(* IEC 61131-3 sources: plc-st-coding-agent/progress/evidence/f14_v14_remaining_20261113/jobs/custom_minimax-m27 (part 5) *)

(* ---- public-medium-05.candidate_04.st ---- *)
(* ENGINEERING_CONTRACT
 * =============================================================================
 * Mode Switching (PUB001): Mode=0 manual, Mode=1 automatic. Output state on
 *   mode transition: both Motor outputs cleared, CompletionLight cleared.
 *   Transition detected via rising edge on Mode input variable.
 * Manual Mode (PUB002/PUB003):
 *   - Activation: Mode=0
 *   - Retention: MotorForward holds while ForwardButton=1 AND ReverseButton=0
 *   - Retention: MotorReverse holds while ReverseButton=1 AND ForwardButton=0
 *   - Deactivation: both cleared on any of: ForwardButton=0, ReverseButton=0,
 *     forward+reverse both asserted (interlock drops both), or Mode→1
 *   - Units: combinational, no timer
 * Automatic Mode (PUB004-PUB008):
 *   - Scan behavior: edge-sensitive state machine evaluated every scan
 *   - STATION_A activation: SensorA=TRUE AND State=IDLE
 *   - STATION_B activation: SensorB=TRUE AND State=MOVING_TO_B
 *   - STATION_C activation: SensorC=TRUE AND State=MOVING_TO_C
 *   - MotorForward activation: (State=IDLE AND SensorA=TRUE→ButtonA=TRUE)
 *     OR (State=STATION_A AND ButtonA=TRUE) OR (State=STATION_B AND ButtonB=TRUE)
 *   - MotorForward deactivation: on SensorB (→STATION_B) or SensorC (→STATION_C)
 *   - CompletionLight activation: SensorC=TRUE AND ButtonC=TRUE AND State=STATION_C
 *   - CompletionLight retention: holds until SensorC=FALSE (product removed)
 *   - CompletionLight deactivation: SensorC=FALSE transitions to IDLE
 *   - IDLE reset: State=IDLE when no product detected at any station
 *   - Units: boolean states, no timers
 * Same-scan priority: manual overrides automatic (Mode check first). Within
 *   automatic, state transition clears prior MotorForward before next sensor
 *   evaluation; CompletionLight set after Mode/state checks finalized.
 * Physical interlock: Pub002 prohibits MotorForward AND MotorReverse together.
 * =============================================================================
 *)

(* CONTRACT_RULES [] *)

FUNCTION_BLOCK ProductionLineControl
VAR_INPUT
    Mode            : BOOL;  (* 0=manual, 1=automatic *)
    ForwardButton   : BOOL;
    ReverseButton   : BOOL;
    SensorA         : BOOL;
    SensorB         : BOOL;
    SensorC         : BOOL;
    ButtonA         : BOOL;
    ButtonB         : BOOL;
    ButtonC         : BOOL;
END_VAR
VAR_OUTPUT
    MotorForward    : BOOL;
    MotorReverse    : BOOL;
    CompletionLight : BOOL;
END_VAR
VAR_CONSTANT
    IDLE         : INT := 0;
    STATION_A    : INT := 1;
    MOVING_TO_B  : INT := 2;
    STATION_B    : INT := 3;
    MOVING_TO_C  : INT := 4;
    STATION_C    : INT := 5;
END_VAR_CONSTANT

VAR
    State           : INT;  (* 0=IDLE, 1=STATION_A, 2=MOVING_TO_B, 3=STATION_B,
                                4=MOVING_TO_C, 5=STATION_C *)
    tmp_PreviousMode : BOOL;
    tmp_ModeRising   : BOOL;
END_VAR

    (* Constants for state identification *)
    (* Detect mode transition for reset behavior *)
    tmp_ModeRising := Mode AND NOT tmp_PreviousMode;
    tmp_PreviousMode := Mode;

    (* Reset outputs on mode entry into automatic *)
    IF tmp_ModeRising THEN
        MotorForward    := FALSE;
        MotorReverse    := FALSE;
        CompletionLight := FALSE;
    END_IF;

    (* Mode-based operation dispatch *)
    IF Mode = FALSE THEN
        (* Manual Mode (PUB002/PUB003) *)
        (* Interlock: forward and reverse cannot be energized together *)
        IF ForwardButton AND NOT ReverseButton THEN
            MotorForward := TRUE;
            MotorReverse := FALSE;
        ELSIF ReverseButton AND NOT ForwardButton THEN
            MotorForward := FALSE;
            MotorReverse := TRUE;
        ELSE
            MotorForward := FALSE;
            MotorReverse := FALSE;
        END_IF;
    ELSE
        (* Automatic Mode (PUB004-PUB008) *)
        MotorForward    := FALSE;
        MotorReverse    := FALSE;

        (* State machine evaluation *)
        CASE State OF
            IDLE :
                (* Wait for product at Workstation A *)
                IF SensorA THEN
                    State := STATION_A;
                END_IF;

            STATION_A :
                (* Product at Workstation A, wait for ButtonA *)
                IF ButtonA THEN
                    MotorForward := TRUE;
                    State := MOVING_TO_B;
                END_IF;
                (* Fallback: if product leaves A unexpectedly, return to IDLE *)
                IF NOT SensorA THEN
                    State := IDLE;
                END_IF;

            MOVING_TO_B :
                (* Motor running forward, wait for SensorB *)
                MotorForward := TRUE;
                IF SensorB THEN
                    MotorForward := FALSE;
                    State := STATION_B;
                END_IF;

            STATION_B :
                (* Product at Workstation B, wait for ButtonB *)
                IF ButtonB THEN
                    MotorForward := TRUE;
                    State := MOVING_TO_C;
                END_IF;
                (* Fallback: if product leaves B unexpectedly, return to IDLE *)
                IF NOT SensorB THEN
                    State := IDLE;
                END_IF;

            MOVING_TO_C :
                (* Motor running forward, wait for SensorC *)
                MotorForward := TRUE;
                IF SensorC THEN
                    MotorForward := FALSE;
                    State := STATION_C;
                END_IF;

            STATION_C :
                (* Product at Workstation C, wait for ButtonC, then product removal *)
                IF ButtonC THEN
                    CompletionLight := TRUE;
                END_IF;
                (* Product taken away: light off, return to IDLE *)
                IF NOT SensorC THEN
                    CompletionLight := FALSE;
                    State := IDLE;
                END_IF;

        END_CASE;
    END_IF;

END_FUNCTION_BLOCK

(* ---- public-medium-05.patch_base_02.st ---- *)
(* ENGINEERING_CONTRACT
 * =============================================================================
 * Mode Switching (PUB001): Mode=0 manual, Mode=1 automatic. Output state on
 *   mode transition: both Motor outputs cleared, CompletionLight cleared.
 *   Transition detected via rising edge on Mode input variable.
 * Manual Mode (PUB002/PUB003):
 *   - Activation: Mode=0
 *   - Retention: MotorForward holds while ForwardButton=1 AND ReverseButton=0
 *   - Retention: MotorReverse holds while ReverseButton=1 AND ForwardButton=0
 *   - Deactivation: both cleared on any of: ForwardButton=0, ReverseButton=0,
 *     forward+reverse both asserted (interlock drops both), or Mode→1
 *   - Units: combinational, no timer
 * Automatic Mode (PUB004-PUB008):
 *   - Scan behavior: edge-sensitive state machine evaluated every scan
 *   - STATION_A activation: SensorA=TRUE AND State=IDLE
 *   - STATION_B activation: SensorB=TRUE AND State=MOVING_TO_B
 *   - STATION_C activation: SensorC=TRUE AND State=MOVING_TO_C
 *   - MotorForward activation: (State=IDLE AND SensorA=TRUE→ButtonA=TRUE)
 *     OR (State=STATION_A AND ButtonA=TRUE) OR (State=STATION_B AND ButtonB=TRUE)
 *   - MotorForward deactivation: on SensorB (→STATION_B) or SensorC (→STATION_C)
 *   - CompletionLight activation: SensorC=TRUE AND ButtonC=TRUE AND State=STATION_C
 *   - CompletionLight retention: holds until SensorC=FALSE (product removed)
 *   - CompletionLight deactivation: SensorC=FALSE transitions to IDLE
 *   - IDLE reset: State=IDLE when no product detected at any station
 *   - Units: boolean states, no timers
 * Same-scan priority: manual overrides automatic (Mode check first). Within
 *   automatic, state transition clears prior MotorForward before next sensor
 *   evaluation; CompletionLight set after Mode/state checks finalized.
 * Physical interlock: Pub002 prohibits MotorForward AND MotorReverse together.
 * =============================================================================
 *)

(* CONTRACT_RULES [] *)

FUNCTION_BLOCK ProductionLineControl
VAR_INPUT
    Mode            : BOOL;  (* 0=manual, 1=automatic *)
    ForwardButton   : BOOL;
    ReverseButton   : BOOL;
    SensorA         : BOOL;
    SensorB         : BOOL;
    SensorC         : BOOL;
    ButtonA         : BOOL;
    ButtonB         : BOOL;
    ButtonC         : BOOL;
END_VAR
VAR_OUTPUT
    MotorForward    : BOOL;
    MotorReverse    : BOOL;
    CompletionLight : BOOL;
END_VAR
VAR
    State           : INT;  (* 0=IDLE, 1=STATION_A, 2=MOVING_TO_B, 3=STATION_B,
                                4=MOVING_TO_C, 5=STATION_C *)
    tmp_PreviousMode : BOOL;
    tmp_ModeRising   : BOOL;
END_VAR

    (* Constants for state identification *)
    CONST
        IDLE         : INT := 0;
        STATION_A    : INT := 1;
        MOVING_TO_B  : INT := 2;
        STATION_B    : INT := 3;
        MOVING_TO_C  : INT := 4;
        STATION_C    : INT := 5;
    END_CONST

    (* Detect mode transition for reset behavior *)
    tmp_ModeRising := Mode AND NOT tmp_PreviousMode;
    tmp_PreviousMode := Mode;

    (* Reset outputs on mode entry into automatic *)
    IF tmp_ModeRising THEN
        MotorForward    := FALSE;
        MotorReverse    := FALSE;
        CompletionLight := FALSE;
    END_IF;

    (* Mode-based operation dispatch *)
    IF Mode = FALSE THEN
        (* Manual Mode (PUB002/PUB003) *)
        (* Interlock: forward and reverse cannot be energized together *)
        IF ForwardButton AND NOT ReverseButton THEN
            MotorForward := TRUE;
            MotorReverse := FALSE;
        ELSIF ReverseButton AND NOT ForwardButton THEN
            MotorForward := FALSE;
            MotorReverse := TRUE;
        ELSE
            MotorForward := FALSE;
            MotorReverse := FALSE;
        END_IF;
    ELSE
        (* Automatic Mode (PUB004-PUB008) *)
        MotorForward    := FALSE;
        MotorReverse    := FALSE;

        (* State machine evaluation *)
        CASE State OF
            IDLE :
                (* Wait for product at Workstation A *)
                IF SensorA THEN
                    State := STATION_A;
                END_IF;

            STATION_A :
                (* Product at Workstation A, wait for ButtonA *)
                IF ButtonA THEN
                    MotorForward := TRUE;
                    State := MOVING_TO_B;
                END_IF;
                (* Fallback: if product leaves A unexpectedly, return to IDLE *)
                IF NOT SensorA THEN
                    State := IDLE;
                END_IF;

            MOVING_TO_B :
                (* Motor running forward, wait for SensorB *)
                MotorForward := TRUE;
                IF SensorB THEN
                    MotorForward := FALSE;
                    State := STATION_B;
                END_IF;

            STATION_B :
                (* Product at Workstation B, wait for ButtonB *)
                IF ButtonB THEN
                    MotorForward := TRUE;
                    State := MOVING_TO_C;
                END_IF;
                (* Fallback: if product leaves B unexpectedly, return to IDLE *)
                IF NOT SensorB THEN
                    State := IDLE;
                END_IF;

            MOVING_TO_C :
                (* Motor running forward, wait for SensorC *)
                MotorForward := TRUE;
                IF SensorC THEN
                    MotorForward := FALSE;
                    State := STATION_C;
                END_IF;

            STATION_C :
                (* Product at Workstation C, wait for ButtonC, then product removal *)
                IF ButtonC THEN
                    CompletionLight := TRUE;
                END_IF;
                (* Product taken away: light off, return to IDLE *)
                IF NOT SensorC THEN
                    CompletionLight := FALSE;
                    State := IDLE;
                END_IF;

        END_CASE;
    END_IF;

END_FUNCTION_BLOCK

(* ---- public-medium-05.patch_base_03.st ---- *)
TYPE ProductionState : INT (
    IDLE := 0,
    STATION_A := 1,
    MOVING_TO_B := 2,
    STATION_B := 3,
    MOVING_TO_C := 4,
    STATION_C := 5
);
END_TYPE;

(* ENGINEERING_CONTRACT
 * =============================================================================
 * Mode Switching (PUB001): Mode=0 manual, Mode=1 automatic. Output state on
 *   mode transition: both Motor outputs cleared, CompletionLight cleared.
 *   Transition detected via rising edge on Mode input variable.
 * Manual Mode (PUB002/PUB003):
 *   - Activation: Mode=0
 *   - Retention: MotorForward holds while ForwardButton=1 AND ReverseButton=0
 *   - Retention: MotorReverse holds while ReverseButton=1 AND ForwardButton=0
 *   - Deactivation: both cleared on any of: ForwardButton=0, ReverseButton=0,
 *     forward+reverse both asserted (interlock drops both), or Mode→1
 *   - Units: combinational, no timer
 * Automatic Mode (PUB004-PUB008):
 *   - Scan behavior: edge-sensitive state machine evaluated every scan
 *   - STATION_A activation: SensorA=TRUE AND State=IDLE
 *   - STATION_B activation: SensorB=TRUE AND State=MOVING_TO_B
 *   - STATION_C activation: SensorC=TRUE AND State=MOVING_TO_C
 *   - MotorForward activation: (State=IDLE AND SensorA=TRUE→ButtonA=TRUE)
 *     OR (State=STATION_A AND ButtonA=TRUE) OR (State=STATION_B AND ButtonB=TRUE)
 *   - MotorForward deactivation: on SensorB (→STATION_B) or SensorC (→STATION_C)
 *   - CompletionLight activation: SensorC=TRUE AND ButtonC=TRUE AND State=STATION_C
 *   - CompletionLight retention: holds until SensorC=FALSE (product removed)
 *   - CompletionLight deactivation: SensorC=FALSE transitions to IDLE
 *   - IDLE reset: State=IDLE when no product detected at any station
 *   - Units: boolean states, no timers
 * Same-scan priority: manual overrides automatic (Mode check first). Within
 *   automatic, state transition clears prior MotorForward before next sensor
 *   evaluation; CompletionLight set after Mode/state checks finalized.
 * Physical interlock: Pub002 prohibits MotorForward AND MotorReverse together.
 * =============================================================================
 *)

(* CONTRACT_RULES [] *)

FUNCTION_BLOCK ProductionLineControl
VAR_INPUT
    Mode            : BOOL;  (* 0=manual, 1=automatic *)
    ForwardButton   : BOOL;
    ReverseButton   : BOOL;
    SensorA         : BOOL;
    SensorB         : BOOL;
    SensorC         : BOOL;
    ButtonA         : BOOL;
    ButtonB         : BOOL;
    ButtonC         : BOOL;
END_VAR
VAR_OUTPUT
    MotorForward    : BOOL;
    MotorReverse    : BOOL;
    CompletionLight : BOOL;
END_VAR
VAR
    State           : INT;  (* 0=IDLE, 1=STATION_A, 2=MOVING_TO_B, 3=STATION_B,
                                4=MOVING_TO_C, 5=STATION_C *)
    tmp_PreviousMode : BOOL;
    tmp_ModeRising   : BOOL;
END_VAR

    (* Constants for state identification *)
    (* Detect mode transition for reset behavior *)
    tmp_ModeRising := Mode AND NOT tmp_PreviousMode;
    tmp_PreviousMode := Mode;

    (* Reset outputs on mode entry into automatic *)
    IF tmp_ModeRising THEN
        MotorForward    := FALSE;
        MotorReverse    := FALSE;
        CompletionLight := FALSE;
    END_IF;

    (* Mode-based operation dispatch *)
    IF Mode = FALSE THEN
        (* Manual Mode (PUB002/PUB003) *)
        (* Interlock: forward and reverse cannot be energized together *)
        IF ForwardButton AND NOT ReverseButton THEN
            MotorForward := TRUE;
            MotorReverse := FALSE;
        ELSIF ReverseButton AND NOT ForwardButton THEN
            MotorForward := FALSE;
            MotorReverse := TRUE;
        ELSE
            MotorForward := FALSE;
            MotorReverse := FALSE;
        END_IF;
    ELSE
        (* Automatic Mode (PUB004-PUB008) *)
        MotorForward    := FALSE;
        MotorReverse    := FALSE;

        (* State machine evaluation *)
        CASE State OF
            IDLE :
                (* Wait for product at Workstation A *)
                IF SensorA THEN
                    State := STATION_A;
                END_IF;

            STATION_A :
                (* Product at Workstation A, wait for ButtonA *)
                IF ButtonA THEN
                    MotorForward := TRUE;
                    State := MOVING_TO_B;
                END_IF;
                (* Fallback: if product leaves A unexpectedly, return to IDLE *)
                IF NOT SensorA THEN
                    State := IDLE;
                END_IF;

            MOVING_TO_B :
                (* Motor running forward, wait for SensorB *)
                MotorForward := TRUE;
                IF SensorB THEN
                    MotorForward := FALSE;
                    State := STATION_B;
                END_IF;

            STATION_B :
                (* Product at Workstation B, wait for ButtonB *)
                IF ButtonB THEN
                    MotorForward := TRUE;
                    State := MOVING_TO_C;
                END_IF;
                (* Fallback: if product leaves B unexpectedly, return to IDLE *)
                IF NOT SensorB THEN
                    State := IDLE;
                END_IF;

            MOVING_TO_C :
                (* Motor running forward, wait for SensorC *)
                MotorForward := TRUE;
                IF SensorC THEN
                    MotorForward := FALSE;
                    State := STATION_C;
                END_IF;

            STATION_C :
                (* Product at Workstation C, wait for ButtonC, then product removal *)
                IF ButtonC THEN
                    CompletionLight := TRUE;
                END_IF;
                (* Product taken away: light off, return to IDLE *)
                IF NOT SensorC THEN
                    CompletionLight := FALSE;
                    State := IDLE;
                END_IF;

        END_CASE;
    END_IF;

END_FUNCTION_BLOCK

(* ---- public-medium-05.patch_base_04.st ---- *)
CONST
    IDLE         : INT := 0;
    STATION_A    : INT := 1;
    MOVING_TO_B  : INT := 2;
    STATION_B    : INT := 3;
    MOVING_TO_C  : INT := 4;
    STATION_C    : INT := 5;
END_CONST

(* ENGINEERING_CONTRACT
 * =============================================================================
 * Mode Switching (PUB001): Mode=0 manual, Mode=1 automatic. Output state on
 *   mode transition: both Motor outputs cleared, CompletionLight cleared.
 *   Transition detected via rising edge on Mode input variable.
 * Manual Mode (PUB002/PUB003):
 *   - Activation: Mode=0
 *   - Retention: MotorForward holds while ForwardButton=1 AND ReverseButton=0
 *   - Retention: MotorReverse holds while ReverseButton=1 AND ForwardButton=0
 *   - Deactivation: both cleared on any of: ForwardButton=0, ReverseButton=0,
 *     forward+reverse both asserted (interlock drops both), or Mode→1
 *   - Units: combinational, no timer
 * Automatic Mode (PUB004-PUB008):
 *   - Scan behavior: edge-sensitive state machine evaluated every scan
 *   - STATION_A activation: SensorA=TRUE AND State=IDLE
 *   - STATION_B activation: SensorB=TRUE AND State=MOVING_TO_B
 *   - STATION_C activation: SensorC=TRUE AND State=MOVING_TO_C
 *   - MotorForward activation: (State=IDLE AND SensorA=TRUE→ButtonA=TRUE)
 *     OR (State=STATION_A AND ButtonA=TRUE) OR (State=STATION_B AND ButtonB=TRUE)
 *   - MotorForward deactivation: on SensorB (→STATION_B) or SensorC (→STATION_C)
 *   - CompletionLight activation: SensorC=TRUE AND ButtonC=TRUE AND State=STATION_C
 *   - CompletionLight retention: holds until SensorC=FALSE (product removed)
 *   - CompletionLight deactivation: SensorC=FALSE transitions to IDLE
 *   - IDLE reset: State=IDLE when no product detected at any station
 *   - Units: boolean states, no timers
 * Same-scan priority: manual overrides automatic (Mode check first). Within
 *   automatic, state transition clears prior MotorForward before next sensor
 *   evaluation; CompletionLight set after Mode/state checks finalized.
 * Physical interlock: Pub002 prohibits MotorForward AND MotorReverse together.
 * =============================================================================
 *)

(* CONTRACT_RULES [] *)

FUNCTION_BLOCK ProductionLineControl
VAR_INPUT
    Mode            : BOOL;  (* 0=manual, 1=automatic *)
    ForwardButton   : BOOL;
    ReverseButton   : BOOL;
    SensorA         : BOOL;
    SensorB         : BOOL;
    SensorC         : BOOL;
    ButtonA         : BOOL;
    ButtonB         : BOOL;
    ButtonC         : BOOL;
END_VAR
VAR_OUTPUT
    MotorForward    : BOOL;
    MotorReverse    : BOOL;
    CompletionLight : BOOL;
END_VAR
VAR
    State           : INT;  (* 0=IDLE, 1=STATION_A, 2=MOVING_TO_B, 3=STATION_B,
                                4=MOVING_TO_C, 5=STATION_C *)
    tmp_PreviousMode : BOOL;
    tmp_ModeRising   : BOOL;
END_VAR

    (* Constants for state identification *)
    (* Detect mode transition for reset behavior *)
    tmp_ModeRising := Mode AND NOT tmp_PreviousMode;
    tmp_PreviousMode := Mode;

    (* Reset outputs on mode entry into automatic *)
    IF tmp_ModeRising THEN
        MotorForward    := FALSE;
        MotorReverse    := FALSE;
        CompletionLight := FALSE;
    END_IF;

    (* Mode-based operation dispatch *)
    IF Mode = FALSE THEN
        (* Manual Mode (PUB002/PUB003) *)
        (* Interlock: forward and reverse cannot be energized together *)
        IF ForwardButton AND NOT ReverseButton THEN
            MotorForward := TRUE;
            MotorReverse := FALSE;
        ELSIF ReverseButton AND NOT ForwardButton THEN
            MotorForward := FALSE;
            MotorReverse := TRUE;
        ELSE
            MotorForward := FALSE;
            MotorReverse := FALSE;
        END_IF;
    ELSE
        (* Automatic Mode (PUB004-PUB008) *)
        MotorForward    := FALSE;
        MotorReverse    := FALSE;

        (* State machine evaluation *)
        CASE State OF
            IDLE :
                (* Wait for product at Workstation A *)
                IF SensorA THEN
                    State := STATION_A;
                END_IF;

            STATION_A :
                (* Product at Workstation A, wait for ButtonA *)
                IF ButtonA THEN
                    MotorForward := TRUE;
                    State := MOVING_TO_B;
                END_IF;
                (* Fallback: if product leaves A unexpectedly, return to IDLE *)
                IF NOT SensorA THEN
                    State := IDLE;
                END_IF;

            MOVING_TO_B :
                (* Motor running forward, wait for SensorB *)
                MotorForward := TRUE;
                IF SensorB THEN
                    MotorForward := FALSE;
                    State := STATION_B;
                END_IF;

            STATION_B :
                (* Product at Workstation B, wait for ButtonB *)
                IF ButtonB THEN
                    MotorForward := TRUE;
                    State := MOVING_TO_C;
                END_IF;
                (* Fallback: if product leaves B unexpectedly, return to IDLE *)
                IF NOT SensorB THEN
                    State := IDLE;
                END_IF;

            MOVING_TO_C :
                (* Motor running forward, wait for SensorC *)
                MotorForward := TRUE;
                IF SensorC THEN
                    MotorForward := FALSE;
                    State := STATION_C;
                END_IF;

            STATION_C :
                (* Product at Workstation C, wait for ButtonC, then product removal *)
                IF ButtonC THEN
                    CompletionLight := TRUE;
                END_IF;
                (* Product taken away: light off, return to IDLE *)
                IF NOT SensorC THEN
                    CompletionLight := FALSE;
                    State := IDLE;
                END_IF;

        END_CASE;
    END_IF;

END_FUNCTION_BLOCK

(* ---- public-medium-05.raw_candidate_01.st ---- *)
(* ENGINEERING_CONTRACT
 * =============================================================================
 * Mode Switching (PUB001): Mode=0 manual, Mode=1 automatic. Output state on
 *   mode transition: both Motor outputs cleared, CompletionLight cleared.
 *   Transition detected via rising edge on Mode input variable.
 * Manual Mode (PUB002/PUB003):
 *   - Activation: Mode=0
 *   - Retention: MotorForward holds while ForwardButton=1 AND ReverseButton=0
 *   - Retention: MotorReverse holds while ReverseButton=1 AND ForwardButton=0
 *   - Deactivation: both cleared on any of: ForwardButton=0, ReverseButton=0,
 *     forward+reverse both asserted (interlock drops both), or Mode→1
 *   - Units: combinational, no timer
 * Automatic Mode (PUB004-PUB008):
 *   - Scan behavior: edge-sensitive state machine evaluated every scan
 *   - STATION_A activation: SensorA=TRUE AND State=IDLE
 *   - STATION_B activation: SensorB=TRUE AND State=MOVING_TO_B
 *   - STATION_C activation: SensorC=TRUE AND State=MOVING_TO_C
 *   - MotorForward activation: (State=IDLE AND SensorA=TRUE→ButtonA=TRUE)
 *     OR (State=STATION_A AND ButtonA=TRUE) OR (State=STATION_B AND ButtonB=TRUE)
 *   - MotorForward deactivation: on SensorB (→STATION_B) or SensorC (→STATION_C)
 *   - CompletionLight activation: SensorC=TRUE AND ButtonC=TRUE AND State=STATION_C
 *   - CompletionLight retention: holds until SensorC=FALSE (product removed)
 *   - CompletionLight deactivation: SensorC=FALSE transitions to IDLE
 *   - IDLE reset: State=IDLE when no product detected at any station
 *   - Units: boolean states, no timers
 * Same-scan priority: manual overrides automatic (Mode check first). Within
 *   automatic, state transition clears prior MotorForward before next sensor
 *   evaluation; CompletionLight set after Mode/state checks finalized.
 * Physical interlock: Pub002 prohibits MotorForward AND MotorReverse together.
 * =============================================================================
 *)

(* CONTRACT_RULES [] *)

FUNCTION_BLOCK ProductionLineControl
VAR_INPUT
    Mode            : BOOL;  (* 0=manual, 1=automatic *)
    ForwardButton   : BOOL;
    ReverseButton   : BOOL;
    SensorA         : BOOL;
    SensorB         : BOOL;
    SensorC         : BOOL;
    ButtonA         : BOOL;
    ButtonB         : BOOL;
    ButtonC         : BOOL;
END_VAR
VAR_OUTPUT
    MotorForward    : BOOL;
    MotorReverse    : BOOL;
    CompletionLight : BOOL;
END_VAR
VAR
    State           : INT;  (* 0=IDLE, 1=STATION_A, 2=MOVING_TO_B, 3=STATION_B,
                                4=MOVING_TO_C, 5=STATION_C *)
    tmp_PreviousMode : BOOL;
    tmp_ModeRising   : BOOL;
END_VAR

    (* Constants for state identification *)
    CONST
        IDLE         : INT := 0;
        STATION_A    : INT := 1;
        MOVING_TO_B  : INT := 2;
        STATION_B    : INT := 3;
        MOVING_TO_C  : INT := 4;
        STATION_C    : INT := 5;
    END_CONST

    (* Detect mode transition for reset behavior *)
    tmp_ModeRising := Mode AND NOT tmp_PreviousMode;
    tmp_PreviousMode := Mode;

    (* Reset outputs on mode entry into automatic *)
    IF tmp_ModeRising THEN
        MotorForward    := FALSE;
        MotorReverse    := FALSE;
        CompletionLight := FALSE;
    END_IF

    (* Mode-based operation dispatch *)
    IF Mode = FALSE THEN
        (* Manual Mode (PUB002/PUB003) *)
        (* Interlock: forward and reverse cannot be energized together *)
        IF ForwardButton AND NOT ReverseButton THEN
            MotorForward := TRUE;
            MotorReverse := FALSE;
        ELSIF ReverseButton AND NOT ForwardButton THEN
            MotorForward := FALSE;
            MotorReverse := TRUE;
        ELSE
            MotorForward := FALSE;
            MotorReverse := FALSE;
        END_IF
    ELSE
        (* Automatic Mode (PUB004-PUB008) *)
        MotorForward    := FALSE;
        MotorReverse    := FALSE;

        (* State machine evaluation *)
        CASE State OF
            IDLE :
                (* Wait for product at Workstation A *)
                IF SensorA THEN
                    State := STATION_A;
                END_IF

            STATION_A :
                (* Product at Workstation A, wait for ButtonA *)
                IF ButtonA THEN
                    MotorForward := TRUE;
                    State := MOVING_TO_B;
                END_IF
                (* Fallback: if product leaves A unexpectedly, return to IDLE *)
                IF NOT SensorA THEN
                    State := IDLE;
                END_IF

            MOVING_TO_B :
                (* Motor running forward, wait for SensorB *)
                MotorForward := TRUE;
                IF SensorB THEN
                    MotorForward := FALSE;
                    State := STATION_B;
                END_IF

            STATION_B :
                (* Product at Workstation B, wait for ButtonB *)
                IF ButtonB THEN
                    MotorForward := TRUE;
                    State := MOVING_TO_C;
                END_IF
                (* Fallback: if product leaves B unexpectedly, return to IDLE *)
                IF NOT SensorB THEN
                    State := IDLE;
                END_IF

            MOVING_TO_C :
                (* Motor running forward, wait for SensorC *)
                MotorForward := TRUE;
                IF SensorC THEN
                    MotorForward := FALSE;
                    State := STATION_C;
                END_IF

            STATION_C :
                (* Product at Workstation C, wait for ButtonC, then product removal *)
                IF ButtonC THEN
                    CompletionLight := TRUE;
                END_IF
                (* Product taken away: light off, return to IDLE *)
                IF NOT SensorC THEN
                    CompletionLight := FALSE;
                    State := IDLE;
                END_IF

        END_CASE
    END_IF

END_FUNCTION_BLOCK

(* ---- public-medium-05.raw_candidate_02.st ---- *)
TYPE ProductionState : INT (
    IDLE := 0,
    STATION_A := 1,
    MOVING_TO_B := 2,
    STATION_B := 3,
    MOVING_TO_C := 4,
    STATION_C := 5
);
END_TYPE

(* ENGINEERING_CONTRACT
 * =============================================================================
 * Mode Switching (PUB001): Mode=0 manual, Mode=1 automatic. Output state on
 *   mode transition: both Motor outputs cleared, CompletionLight cleared.
 *   Transition detected via rising edge on Mode input variable.
 * Manual Mode (PUB002/PUB003):
 *   - Activation: Mode=0
 *   - Retention: MotorForward holds while ForwardButton=1 AND ReverseButton=0
 *   - Retention: MotorReverse holds while ReverseButton=1 AND ForwardButton=0
 *   - Deactivation: both cleared on any of: ForwardButton=0, ReverseButton=0,
 *     forward+reverse both asserted (interlock drops both), or Mode→1
 *   - Units: combinational, no timer
 * Automatic Mode (PUB004-PUB008):
 *   - Scan behavior: edge-sensitive state machine evaluated every scan
 *   - STATION_A activation: SensorA=TRUE AND State=IDLE
 *   - STATION_B activation: SensorB=TRUE AND State=MOVING_TO_B
 *   - STATION_C activation: SensorC=TRUE AND State=MOVING_TO_C
 *   - MotorForward activation: (State=IDLE AND SensorA=TRUE→ButtonA=TRUE)
 *     OR (State=STATION_A AND ButtonA=TRUE) OR (State=STATION_B AND ButtonB=TRUE)
 *   - MotorForward deactivation: on SensorB (→STATION_B) or SensorC (→STATION_C)
 *   - CompletionLight activation: SensorC=TRUE AND ButtonC=TRUE AND State=STATION_C
 *   - CompletionLight retention: holds until SensorC=FALSE (product removed)
 *   - CompletionLight deactivation: SensorC=FALSE transitions to IDLE
 *   - IDLE reset: State=IDLE when no product detected at any station
 *   - Units: boolean states, no timers
 * Same-scan priority: manual overrides automatic (Mode check first). Within
 *   automatic, state transition clears prior MotorForward before next sensor
 *   evaluation; CompletionLight set after Mode/state checks finalized.
 * Physical interlock: Pub002 prohibits MotorForward AND MotorReverse together.
 * =============================================================================
 *)

(* CONTRACT_RULES [] *)

FUNCTION_BLOCK ProductionLineControl
VAR_INPUT
    Mode            : BOOL;  (* 0=manual, 1=automatic *)
    ForwardButton   : BOOL;
    ReverseButton   : BOOL;
    SensorA         : BOOL;
    SensorB         : BOOL;
    SensorC         : BOOL;
    ButtonA         : BOOL;
    ButtonB         : BOOL;
    ButtonC         : BOOL;
END_VAR
VAR_OUTPUT
    MotorForward    : BOOL;
    MotorReverse    : BOOL;
    CompletionLight : BOOL;
END_VAR
VAR
    State           : INT;  (* 0=IDLE, 1=STATION_A, 2=MOVING_TO_B, 3=STATION_B,
                                4=MOVING_TO_C, 5=STATION_C *)
    tmp_PreviousMode : BOOL;
    tmp_ModeRising   : BOOL;
END_VAR

    (* Constants for state identification *)
    (* Detect mode transition for reset behavior *)
    tmp_ModeRising := Mode AND NOT tmp_PreviousMode;
    tmp_PreviousMode := Mode;

    (* Reset outputs on mode entry into automatic *)
    IF tmp_ModeRising THEN
        MotorForward    := FALSE;
        MotorReverse    := FALSE;
        CompletionLight := FALSE;
    END_IF;

    (* Mode-based operation dispatch *)
    IF Mode = FALSE THEN
        (* Manual Mode (PUB002/PUB003) *)
        (* Interlock: forward and reverse cannot be energized together *)
        IF ForwardButton AND NOT ReverseButton THEN
            MotorForward := TRUE;
            MotorReverse := FALSE;
        ELSIF ReverseButton AND NOT ForwardButton THEN
            MotorForward := FALSE;
            MotorReverse := TRUE;
        ELSE
            MotorForward := FALSE;
            MotorReverse := FALSE;
        END_IF;
    ELSE
        (* Automatic Mode (PUB004-PUB008) *)
        MotorForward    := FALSE;
        MotorReverse    := FALSE;

        (* State machine evaluation *)
        CASE State OF
            IDLE :
                (* Wait for product at Workstation A *)
                IF SensorA THEN
                    State := STATION_A;
                END_IF;

            STATION_A :
                (* Product at Workstation A, wait for ButtonA *)
                IF ButtonA THEN
                    MotorForward := TRUE;
                    State := MOVING_TO_B;
                END_IF;
                (* Fallback: if product leaves A unexpectedly, return to IDLE *)
                IF NOT SensorA THEN
                    State := IDLE;
                END_IF;

            MOVING_TO_B :
                (* Motor running forward, wait for SensorB *)
                MotorForward := TRUE;
                IF SensorB THEN
                    MotorForward := FALSE;
                    State := STATION_B;
                END_IF;

            STATION_B :
                (* Product at Workstation B, wait for ButtonB *)
                IF ButtonB THEN
                    MotorForward := TRUE;
                    State := MOVING_TO_C;
                END_IF;
                (* Fallback: if product leaves B unexpectedly, return to IDLE *)
                IF NOT SensorB THEN
                    State := IDLE;
                END_IF;

            MOVING_TO_C :
                (* Motor running forward, wait for SensorC *)
                MotorForward := TRUE;
                IF SensorC THEN
                    MotorForward := FALSE;
                    State := STATION_C;
                END_IF;

            STATION_C :
                (* Product at Workstation C, wait for ButtonC, then product removal *)
                IF ButtonC THEN
                    CompletionLight := TRUE;
                END_IF;
                (* Product taken away: light off, return to IDLE *)
                IF NOT SensorC THEN
                    CompletionLight := FALSE;
                    State := IDLE;
                END_IF;

        END_CASE;
    END_IF;

END_FUNCTION_BLOCK

(* ---- public-medium-05.raw_candidate_03.st ---- *)
CONST
    IDLE         : INT := 0;
    STATION_A    : INT := 1;
    MOVING_TO_B  : INT := 2;
    STATION_B    : INT := 3;
    MOVING_TO_C  : INT := 4;
    STATION_C    : INT := 5;
END_CONST

(* ENGINEERING_CONTRACT
 * =============================================================================
 * Mode Switching (PUB001): Mode=0 manual, Mode=1 automatic. Output state on
 *   mode transition: both Motor outputs cleared, CompletionLight cleared.
 *   Transition detected via rising edge on Mode input variable.
 * Manual Mode (PUB002/PUB003):
 *   - Activation: Mode=0
 *   - Retention: MotorForward holds while ForwardButton=1 AND ReverseButton=0
 *   - Retention: MotorReverse holds while ReverseButton=1 AND ForwardButton=0
 *   - Deactivation: both cleared on any of: ForwardButton=0, ReverseButton=0,
 *     forward+reverse both asserted (interlock drops both), or Mode→1
 *   - Units: combinational, no timer
 * Automatic Mode (PUB004-PUB008):
 *   - Scan behavior: edge-sensitive state machine evaluated every scan
 *   - STATION_A activation: SensorA=TRUE AND State=IDLE
 *   - STATION_B activation: SensorB=TRUE AND State=MOVING_TO_B
 *   - STATION_C activation: SensorC=TRUE AND State=MOVING_TO_C
 *   - MotorForward activation: (State=IDLE AND SensorA=TRUE→ButtonA=TRUE)
 *     OR (State=STATION_A AND ButtonA=TRUE) OR (State=STATION_B AND ButtonB=TRUE)
 *   - MotorForward deactivation: on SensorB (→STATION_B) or SensorC (→STATION_C)
 *   - CompletionLight activation: SensorC=TRUE AND ButtonC=TRUE AND State=STATION_C
 *   - CompletionLight retention: holds until SensorC=FALSE (product removed)
 *   - CompletionLight deactivation: SensorC=FALSE transitions to IDLE
 *   - IDLE reset: State=IDLE when no product detected at any station
 *   - Units: boolean states, no timers
 * Same-scan priority: manual overrides automatic (Mode check first). Within
 *   automatic, state transition clears prior MotorForward before next sensor
 *   evaluation; CompletionLight set after Mode/state checks finalized.
 * Physical interlock: Pub002 prohibits MotorForward AND MotorReverse together.
 * =============================================================================
 *)

(* CONTRACT_RULES [] *)

FUNCTION_BLOCK ProductionLineControl
VAR_INPUT
    Mode            : BOOL;  (* 0=manual, 1=automatic *)
    ForwardButton   : BOOL;
    ReverseButton   : BOOL;
    SensorA         : BOOL;
    SensorB         : BOOL;
    SensorC         : BOOL;
    ButtonA         : BOOL;
    ButtonB         : BOOL;
    ButtonC         : BOOL;
END_VAR
VAR_OUTPUT
    MotorForward    : BOOL;
    MotorReverse    : BOOL;
    CompletionLight : BOOL;
END_VAR
VAR
    State           : INT;  (* 0=IDLE, 1=STATION_A, 2=MOVING_TO_B, 3=STATION_B,
                                4=MOVING_TO_C, 5=STATION_C *)
    tmp_PreviousMode : BOOL;
    tmp_ModeRising   : BOOL;
END_VAR

    (* Constants for state identification *)
    (* Detect mode transition for reset behavior *)
    tmp_ModeRising := Mode AND NOT tmp_PreviousMode;
    tmp_PreviousMode := Mode;

    (* Reset outputs on mode entry into automatic *)
    IF tmp_ModeRising THEN
        MotorForward    := FALSE;
        MotorReverse    := FALSE;
        CompletionLight := FALSE;
    END_IF;

    (* Mode-based operation dispatch *)
    IF Mode = FALSE THEN
        (* Manual Mode (PUB002/PUB003) *)
        (* Interlock: forward and reverse cannot be energized together *)
        IF ForwardButton AND NOT ReverseButton THEN
            MotorForward := TRUE;
            MotorReverse := FALSE;
        ELSIF ReverseButton AND NOT ForwardButton THEN
            MotorForward := FALSE;
            MotorReverse := TRUE;
        ELSE
            MotorForward := FALSE;
            MotorReverse := FALSE;
        END_IF;
    ELSE
        (* Automatic Mode (PUB004-PUB008) *)
        MotorForward    := FALSE;
        MotorReverse    := FALSE;

        (* State machine evaluation *)
        CASE State OF
            IDLE :
                (* Wait for product at Workstation A *)
                IF SensorA THEN
                    State := STATION_A;
                END_IF;

            STATION_A :
                (* Product at Workstation A, wait for ButtonA *)
                IF ButtonA THEN
                    MotorForward := TRUE;
                    State := MOVING_TO_B;
                END_IF;
                (* Fallback: if product leaves A unexpectedly, return to IDLE *)
                IF NOT SensorA THEN
                    State := IDLE;
                END_IF;

            MOVING_TO_B :
                (* Motor running forward, wait for SensorB *)
                MotorForward := TRUE;
                IF SensorB THEN
                    MotorForward := FALSE;
                    State := STATION_B;
                END_IF;

            STATION_B :
                (* Product at Workstation B, wait for ButtonB *)
                IF ButtonB THEN
                    MotorForward := TRUE;
                    State := MOVING_TO_C;
                END_IF;
                (* Fallback: if product leaves B unexpectedly, return to IDLE *)
                IF NOT SensorB THEN
                    State := IDLE;
                END_IF;

            MOVING_TO_C :
                (* Motor running forward, wait for SensorC *)
                MotorForward := TRUE;
                IF SensorC THEN
                    MotorForward := FALSE;
                    State := STATION_C;
                END_IF;

            STATION_C :
                (* Product at Workstation C, wait for ButtonC, then product removal *)
                IF ButtonC THEN
                    CompletionLight := TRUE;
                END_IF;
                (* Product taken away: light off, return to IDLE *)
                IF NOT SensorC THEN
                    CompletionLight := FALSE;
                    State := IDLE;
                END_IF;

        END_CASE;
    END_IF;

END_FUNCTION_BLOCK

(* ---- public-medium-05.raw_candidate_04.st ---- *)
(* ENGINEERING_CONTRACT
 * =============================================================================
 * Mode Switching (PUB001): Mode=0 manual, Mode=1 automatic. Output state on
 *   mode transition: both Motor outputs cleared, CompletionLight cleared.
 *   Transition detected via rising edge on Mode input variable.
 * Manual Mode (PUB002/PUB003):
 *   - Activation: Mode=0
 *   - Retention: MotorForward holds while ForwardButton=1 AND ReverseButton=0
 *   - Retention: MotorReverse holds while ReverseButton=1 AND ForwardButton=0
 *   - Deactivation: both cleared on any of: ForwardButton=0, ReverseButton=0,
 *     forward+reverse both asserted (interlock drops both), or Mode→1
 *   - Units: combinational, no timer
 * Automatic Mode (PUB004-PUB008):
 *   - Scan behavior: edge-sensitive state machine evaluated every scan
 *   - STATION_A activation: SensorA=TRUE AND State=IDLE
 *   - STATION_B activation: SensorB=TRUE AND State=MOVING_TO_B
 *   - STATION_C activation: SensorC=TRUE AND State=MOVING_TO_C
 *   - MotorForward activation: (State=IDLE AND SensorA=TRUE→ButtonA=TRUE)
 *     OR (State=STATION_A AND ButtonA=TRUE) OR (State=STATION_B AND ButtonB=TRUE)
 *   - MotorForward deactivation: on SensorB (→STATION_B) or SensorC (→STATION_C)
 *   - CompletionLight activation: SensorC=TRUE AND ButtonC=TRUE AND State=STATION_C
 *   - CompletionLight retention: holds until SensorC=FALSE (product removed)
 *   - CompletionLight deactivation: SensorC=FALSE transitions to IDLE
 *   - IDLE reset: State=IDLE when no product detected at any station
 *   - Units: boolean states, no timers
 * Same-scan priority: manual overrides automatic (Mode check first). Within
 *   automatic, state transition clears prior MotorForward before next sensor
 *   evaluation; CompletionLight set after Mode/state checks finalized.
 * Physical interlock: Pub002 prohibits MotorForward AND MotorReverse together.
 * =============================================================================
 *)

(* CONTRACT_RULES [] *)

FUNCTION_BLOCK ProductionLineControl
VAR_INPUT
    Mode            : BOOL;  (* 0=manual, 1=automatic *)
    ForwardButton   : BOOL;
    ReverseButton   : BOOL;
    SensorA         : BOOL;
    SensorB         : BOOL;
    SensorC         : BOOL;
    ButtonA         : BOOL;
    ButtonB         : BOOL;
    ButtonC         : BOOL;
END_VAR
VAR_OUTPUT
    MotorForward    : BOOL;
    MotorReverse    : BOOL;
    CompletionLight : BOOL;
END_VAR
VAR_CONSTANT
    IDLE         : INT := 0;
    STATION_A    : INT := 1;
    MOVING_TO_B  : INT := 2;
    STATION_B    : INT := 3;
    MOVING_TO_C  : INT := 4;
    STATION_C    : INT := 5;
END_VAR_CONSTANT

VAR
    State           : INT;  (* 0=IDLE, 1=STATION_A, 2=MOVING_TO_B, 3=STATION_B,
                                4=MOVING_TO_C, 5=STATION_C *)
    tmp_PreviousMode : BOOL;
    tmp_ModeRising   : BOOL;
END_VAR

    (* Constants for state identification *)
    (* Detect mode transition for reset behavior *)
    tmp_ModeRising := Mode AND NOT tmp_PreviousMode;
    tmp_PreviousMode := Mode;

    (* Reset outputs on mode entry into automatic *)
    IF tmp_ModeRising THEN
        MotorForward    := FALSE;
        MotorReverse    := FALSE;
        CompletionLight := FALSE;
    END_IF;

    (* Mode-based operation dispatch *)
    IF Mode = FALSE THEN
        (* Manual Mode (PUB002/PUB003) *)
        (* Interlock: forward and reverse cannot be energized together *)
        IF ForwardButton AND NOT ReverseButton THEN
            MotorForward := TRUE;
            MotorReverse := FALSE;
        ELSIF ReverseButton AND NOT ForwardButton THEN
            MotorForward := FALSE;
            MotorReverse := TRUE;
        ELSE
            MotorForward := FALSE;
            MotorReverse := FALSE;
        END_IF;
    ELSE
        (* Automatic Mode (PUB004-PUB008) *)
        MotorForward    := FALSE;
        MotorReverse    := FALSE;

        (* State machine evaluation *)
        CASE State OF
            IDLE :
                (* Wait for product at Workstation A *)
                IF SensorA THEN
                    State := STATION_A;
                END_IF;

            STATION_A :
                (* Product at Workstation A, wait for ButtonA *)
                IF ButtonA THEN
                    MotorForward := TRUE;
                    State := MOVING_TO_B;
                END_IF;
                (* Fallback: if product leaves A unexpectedly, return to IDLE *)
                IF NOT SensorA THEN
                    State := IDLE;
                END_IF;

            MOVING_TO_B :
                (* Motor running forward, wait for SensorB *)
                MotorForward := TRUE;
                IF SensorB THEN
                    MotorForward := FALSE;
                    State := STATION_B;
                END_IF;

            STATION_B :
                (* Product at Workstation B, wait for ButtonB *)
                IF ButtonB THEN
                    MotorForward := TRUE;
                    State := MOVING_TO_C;
                END_IF;
                (* Fallback: if product leaves B unexpectedly, return to IDLE *)
                IF NOT SensorB THEN
                    State := IDLE;
                END_IF;

            MOVING_TO_C :
                (* Motor running forward, wait for SensorC *)
                MotorForward := TRUE;
                IF SensorC THEN
                    MotorForward := FALSE;
                    State := STATION_C;
                END_IF;

            STATION_C :
                (* Product at Workstation C, wait for ButtonC, then product removal *)
                IF ButtonC THEN
                    CompletionLight := TRUE;
                END_IF;
                (* Product taken away: light off, return to IDLE *)
                IF NOT SensorC THEN
                    CompletionLight := FALSE;
                    State := IDLE;
                END_IF;

        END_CASE;
    END_IF;

END_FUNCTION_BLOCK

(* ---- public-medium-06.candidate_01.st ---- *)
FUNCTION_BLOCK FB_SlabThicknessMonitor
(*
 * ENGINEERING_CONTRACT
 * =============================================================================
 * Output/State          | Activation          | Retention            | Reset/Deactivation            | Units
 * ----------------------+---------------------+----------------------+-------------------------------+-----------------
 * THICKNESS_ALARM       | Rising edge valid   | Min 500ms hold;      | Signal invalid clears all     | BOOL
 *                       | THICKNESS_FAULT     | continues if fault   | alarm and hold state (PUB001) |
 * Alarm hold timer      | TON(IN: valid &     | TON.ET saturates at  | Signal invalid resets TON     | LTIME (≥500ms)
 *                       |   (fault OR holding))| PT=500ms            |                               |
 * Holding flag          | Fault OR holding    | Self-holds while     | Signal invalid clears         | BOOL
 *                       |                     |   fault OR timer run |                               |
 * Slab_Fault_Counter    | FALSE→TRUE valid    | Accumulates monoton  | None by task spec             | UINT
 *                       | fault transition    | (never auto-reset)   |                               |
 * Slab_Fault_History[0] | New fault entry     | Shifts [n]→[n+1]     | Power-up init to 0            | ARRAY[0..4] DINT
 *                       | writes to index 0   | (0 newest)           |                               |
 * Slab_Runtime_Accumulator| While CUTTING_RUN  | Preserved when       | None by task spec             | LTIME (accumulates)
 *                       | + valid + no fault  | conditions not met   |                               |
 * =============================================================================
 * CONTRACT_RULES [{"kind": "hold_until_reset", "output": "THICKNESS_ALARM", "set_input": "THICKNESS_FAULT", "reset_input": null}]
 *)

VAR_INPUT
    THICKNESS_FAULT        : BOOL;
    THICKNESS_SIGNAL_VALID : BOOL;
    CUTTING_RUN            : BOOL;
    FaultTimestamp         : DINT;
    CycleTime              : TIME;
END_VAR

VAR_OUTPUT
    THICKNESS_ALARM           : BOOL;
    Slab_Fault_Counter        : UINT;
    Slab_Runtime_Accumulator  : LTIME;
    Slab_Fault_History        : ARRAY[0..4] OF DINT;
END_VAR

VAR
    faultRisingEdge    : R_TRIG;
    signalValidPrev    : BOOL;
    alarmHoldTimer     : TON;
    alarmHolding       : BOOL;
    faultActive        : BOOL;
END_VAR

// ---------------------------------------------------------------------------
// Power-up initialization (first scan after instantiation)
// ---------------------------------------------------------------------------
IF NOT alarmHoldTimer.Q AND NOT faultActive AND NOT alarmHolding THEN
    Slab_Fault_Counter       := 0;
    Slab_Runtime_Accumulator := LTIME#0s;
    Slab_Fault_History[0]    := 0;
    Slab_Fault_History[1]    := 0;
    Slab_Fault_History[2]    := 0;
    Slab_Fault_History[3]    := 0;
    Slab_Fault_History[4]    := 0;
END_IF;

// ---------------------------------------------------------------------------
// Detect FALSE→TRUE transition on valid fault signal
// ---------------------------------------------------------------------------
faultRisingEdge(CLK := THICKNESS_FAULT AND THICKNESS_SIGNAL_VALID);

// ---------------------------------------------------------------------------
// Handle signal-valid transitions: clear alarm/hold when signal lost (PUB001)
// ---------------------------------------------------------------------------
IF THICKNESS_SIGNAL_VALID THEN
    IF NOT signalValidPrev THEN
        // Signal just restored after being invalid
        alarmHolding  := FALSE;
        alarmHoldTimer(IN := FALSE);
        faultActive   := FALSE;
    END_IF;

    // -------------------------------------------------------------------------
    // On rising edge of valid fault: record entry and start hold
    // -------------------------------------------------------------------------
    IF faultRisingEdge.Q THEN
        // Increment counter
        Slab_Fault_Counter := Slab_Fault_Counter + UINT#1;

        // Shift history: index 3→4, 2→3, 1→2, 0→1, then write new to 0
        Slab_Fault_History[4] := Slab_Fault_History[3];
        Slab_Fault_History[3] := Slab_Fault_History[2];
        Slab_Fault_History[2] := Slab_Fault_History[1];
        Slab_Fault_History[1] := Slab_Fault_History[0];
        Slab_Fault_History[0] := FaultTimestamp;

        // Activate alarm and start 500 ms hold timer
        faultActive        := TRUE;
        alarmHolding       := TRUE;
        alarmHoldTimer(IN  := TRUE, PT := T#500ms);
    END_IF;

    // -------------------------------------------------------------------------
    // Update alarm state: hold while fault persists or timer running
    // -------------------------------------------------------------------------
    IF faultActive THEN
        // Keep timer running while fault is present
        alarmHoldTimer(IN := TRUE, PT := T#500ms);

        // Alarm stays active while fault or hold timer active
        alarmHolding := THICKNESS_FAULT OR alarmHoldTimer.Q;

        // Release hold tracking once fault clears and timer completes
        IF NOT THICKNESS_FAULT AND alarmHolding AND NOT alarmHoldTimer.Q THEN
            alarmHolding := FALSE;
        END_IF;

        // Clear fault-active flag when fault goes away (hold may continue)
        IF NOT THICKNESS_FAULT THEN
            faultActive := FALSE;
        END_IF;
    END_IF;

    // Final alarm output
    THICKNESS_ALARM := alarmHolding OR faultActive;

    // -------------------------------------------------------------------------
    // Runtime accumulation: only while cutting, signal valid, no fault
    // -------------------------------------------------------------------------
    IF CUTTING_RUN AND NOT THICKNESS_FAULT THEN
        Slab_Runtime_Accumulator := Slab_Runtime_Accumulator + CycleTime;
    END_IF;

ELSE
    // Signal invalid: clear alarm and all hold state (PUB001)
    THICKNESS_ALARM  := FALSE;
    alarmHolding     := FALSE;
    faultActive      := FALSE;
    alarmHoldTimer(IN := FALSE);
END_IF;

// ---------------------------------------------------------------------------
// Latch previous scan signal-valid state for edge detection
// ---------------------------------------------------------------------------
signalValidPrev := THICKNESS_SIGNAL_VALID;

END_FUNCTION_BLOCK

(* ---- public-medium-06.candidate_02.st ---- *)
FUNCTION_BLOCK FB_SlabThicknessMonitor
(*
 * ENGINEERING_CONTRACT
 * =============================================================================
 * Output/State          | Activation          | Retention            | Reset/Deactivation            | Units
 * ----------------------+---------------------+----------------------+-------------------------------+-----------------
 * THICKNESS_ALARM       | Rising edge valid   | Min 500ms hold;      | Signal invalid clears all     | BOOL
 *                       | THICKNESS_FAULT     | continues if fault   | alarm and hold state (PUB001) |
 * Alarm hold timer      | TON(IN: valid &     | TON.ET saturates at  | Signal invalid resets TON     | LTIME (≥500ms)
 *                       |   (fault OR holding))| PT=500ms            |                               |
 * Holding flag          | Fault OR holding    | Self-holds while     | Signal invalid clears         | BOOL
 *                       |                     |   fault OR timer run |                               |
 * Slab_Fault_Counter    | FALSE→TRUE valid    | Accumulates monoton  | None by task spec             | UINT
 *                       | fault transition    | (never auto-reset)   |                               |
 * Slab_Fault_History[0] | New fault entry     | Shifts [n]→[n+1]     | Power-up init to 0            | ARRAY[0..4] DINT
 *                       | writes to index 0   | (0 newest)           |                               |
 * Slab_Runtime_Accumulator| While CUTTING_RUN  | Preserved when       | None by task spec             | LTIME (accumulates)
 *                       | + valid + no fault  | conditions not met   |                               |
 * =============================================================================
 * CONTRACT_RULES [{"kind": "hold_until_reset", "output": "THICKNESS_ALARM", "set_input": "THICKNESS_FAULT", "reset_input": null}]
 *)

VAR_INPUT
    THICKNESS_FAULT        : BOOL;
    THICKNESS_SIGNAL_VALID : BOOL;
    CUTTING_RUN            : BOOL;
    FaultTimestamp         : DINT;
    CycleTime              : TIME;
END_VAR

VAR_OUTPUT
    THICKNESS_ALARM           : BOOL;
    Slab_Fault_Counter        : UINT;
    Slab_Runtime_Accumulator  : LTIME;
    Slab_Fault_History        : ARRAY[0..4] OF DINT;
END_VAR

VAR
    faultRisingEdge    : R_TRIG;
    signalValidPrev    : BOOL;
    alarmHoldTimer     : TON;
    alarmHolding       : BOOL;
    faultActive        : BOOL;
END_VAR

// ---------------------------------------------------------------------------
// Power-up initialization (first scan after instantiation)
// ---------------------------------------------------------------------------
IF NOT alarmHoldTimer.Q AND NOT faultActive AND NOT alarmHolding THEN
    Slab_Fault_Counter       := 0;
    Slab_Runtime_Accumulator := LTIME#0;
    Slab_Fault_History[0]    := 0;
    Slab_Fault_History[1]    := 0;
    Slab_Fault_History[2]    := 0;
    Slab_Fault_History[3]    := 0;
    Slab_Fault_History[4]    := 0;
END_IF;

// ---------------------------------------------------------------------------
// Detect FALSE→TRUE transition on valid fault signal
// ---------------------------------------------------------------------------
faultRisingEdge(CLK := THICKNESS_FAULT AND THICKNESS_SIGNAL_VALID);

// ---------------------------------------------------------------------------
// Handle signal-valid transitions: clear alarm/hold when signal lost (PUB001)
// ---------------------------------------------------------------------------
IF THICKNESS_SIGNAL_VALID THEN
    IF NOT signalValidPrev THEN
        // Signal just restored after being invalid
        alarmHolding  := FALSE;
        alarmHoldTimer(IN := FALSE);
        faultActive   := FALSE;
    END_IF;

    // -------------------------------------------------------------------------
    // On rising edge of valid fault: record entry and start hold
    // -------------------------------------------------------------------------
    IF faultRisingEdge.Q THEN
        // Increment counter
        Slab_Fault_Counter := Slab_Fault_Counter + UINT#1;

        // Shift history: index 3→4, 2→3, 1→2, 0→1, then write new to 0
        Slab_Fault_History[4] := Slab_Fault_History[3];
        Slab_Fault_History[3] := Slab_Fault_History[2];
        Slab_Fault_History[2] := Slab_Fault_History[1];
        Slab_Fault_History[1] := Slab_Fault_History[0];
        Slab_Fault_History[0] := FaultTimestamp;

        // Activate alarm and start 500 ms hold timer
        faultActive        := TRUE;
        alarmHolding       := TRUE;
        alarmHoldTimer(IN  := TRUE, PT := T#500ms);
    END_IF;

    // -------------------------------------------------------------------------
    // Update alarm state: hold while fault persists or timer running
    // -------------------------------------------------------------------------
    IF faultActive THEN
        // Keep timer running while fault is present
        alarmHoldTimer(IN := TRUE, PT := T#500ms);

        // Alarm stays active while fault or hold timer active
        alarmHolding := THICKNESS_FAULT OR alarmHoldTimer.Q;

        // Release hold tracking once fault clears and timer completes
        IF NOT THICKNESS_FAULT AND alarmHolding AND NOT alarmHoldTimer.Q THEN
            alarmHolding := FALSE;
        END_IF;

        // Clear fault-active flag when fault goes away (hold may continue)
        IF NOT THICKNESS_FAULT THEN
            faultActive := FALSE;
        END_IF;
    END_IF;

    // Final alarm output
    THICKNESS_ALARM := alarmHolding OR faultActive;

    // -------------------------------------------------------------------------
    // Runtime accumulation: only while cutting, signal valid, no fault
    // -------------------------------------------------------------------------
    IF CUTTING_RUN AND NOT THICKNESS_FAULT THEN
        Slab_Runtime_Accumulator := Slab_Runtime_Accumulator + TO_LTIME(CycleTime);
    END_IF;

ELSE
    // Signal invalid: clear alarm and all hold state (PUB001)
    THICKNESS_ALARM  := FALSE;
    alarmHolding     := FALSE;
    faultActive      := FALSE;
    alarmHoldTimer(IN := FALSE);
END_IF;

// ---------------------------------------------------------------------------
// Latch previous scan signal-valid state for edge detection
// ---------------------------------------------------------------------------
signalValidPrev := THICKNESS_SIGNAL_VALID;

END_FUNCTION_BLOCK

(* ---- public-medium-06.candidate_03.st ---- *)
FUNCTION_BLOCK FB_SlabThicknessMonitor
(*
 * ENGINEERING_CONTRACT
 * =============================================================================
 * Output/State          | Activation          | Retention            | Reset/Deactivation            | Units
 * ----------------------+---------------------+----------------------+-------------------------------+-----------------
 * THICKNESS_ALARM       | Rising edge valid   | Min 500ms hold;      | Signal invalid clears all     | BOOL
 *                       | THICKNESS_FAULT     | continues if fault   | alarm and hold state (PUB001) |
 * Alarm hold timer      | TON(IN: valid &     | TON.ET saturates at  | Signal invalid resets TON     | LTIME (≥500ms)
 *                       |   (fault OR holding))| PT=500ms            |                               |
 * Holding flag          | Fault OR holding    | Self-holds while     | Signal invalid clears         | BOOL
 *                       |                     |   fault OR timer run |                               |
 * Slab_Fault_Counter    | FALSE→TRUE valid    | Accumulates monoton  | None by task spec             | UINT
 *                       | fault transition    | (never auto-reset)   |                               |
 * Slab_Fault_History[0] | New fault entry     | Shifts [n]→[n+1]     | Power-up init to 0            | ARRAY[0..4] DINT
 *                       | writes to index 0   | (0 newest)           |                               |
 * Slab_Runtime_Accumulator| While CUTTING_RUN  | Preserved when       | None by task spec             | LTIME (accumulates)
 *                       | + valid + no fault  | conditions not met   |                               |
 * =============================================================================
 * CONTRACT_RULES [{"kind": "hold_until_reset", "output": "THICKNESS_ALARM", "set_input": "THICKNESS_FAULT", "reset_input": null}]
 *)

VAR_INPUT
    THICKNESS_FAULT        : BOOL;
    THICKNESS_SIGNAL_VALID : BOOL;
    CUTTING_RUN            : BOOL;
    FaultTimestamp         : DINT;
    CycleTime              : TIME;
END_VAR

VAR_OUTPUT
    THICKNESS_ALARM           : BOOL;
    Slab_Fault_Counter        : UINT;
    Slab_Runtime_Accumulator  : LTIME;
    Slab_Fault_History        : ARRAY[0..4] OF DINT;
END_VAR

VAR
    faultRisingEdge    : R_TRIG;
    signalValidPrev    : BOOL;
    alarmHoldTimer     : TON;
    alarmHolding       : BOOL;
    faultActive        : BOOL;
END_VAR

// ---------------------------------------------------------------------------
// Power-up initialization (first scan after instantiation)
// ---------------------------------------------------------------------------
IF NOT alarmHoldTimer.Q AND NOT faultActive AND NOT alarmHolding THEN
    Slab_Fault_Counter       := 0;
    Slab_Runtime_Accumulator := LTIME#0ms;
    Slab_Fault_History[0]    := 0;
    Slab_Fault_History[1]    := 0;
    Slab_Fault_History[2]    := 0;
    Slab_Fault_History[3]    := 0;
    Slab_Fault_History[4]    := 0;
END_IF;

// ---------------------------------------------------------------------------
// Detect FALSE→TRUE transition on valid fault signal
// ---------------------------------------------------------------------------
faultRisingEdge(CLK := THICKNESS_FAULT AND THICKNESS_SIGNAL_VALID);

// ---------------------------------------------------------------------------
// Handle signal-valid transitions: clear alarm/hold when signal lost (PUB001)
// ---------------------------------------------------------------------------
IF THICKNESS_SIGNAL_VALID THEN
    IF NOT signalValidPrev THEN
        // Signal just restored after being invalid
        alarmHolding  := FALSE;
        alarmHoldTimer(IN := FALSE);
        faultActive   := FALSE;
    END_IF;

    // -------------------------------------------------------------------------
    // On rising edge of valid fault: record entry and start hold
    // -------------------------------------------------------------------------
    IF faultRisingEdge.Q THEN
        // Increment counter
        Slab_Fault_Counter := Slab_Fault_Counter + UINT#1;

        // Shift history: index 3→4, 2→3, 1→2, 0→1, then write new to 0
        Slab_Fault_History[4] := Slab_Fault_History[3];
        Slab_Fault_History[3] := Slab_Fault_History[2];
        Slab_Fault_History[2] := Slab_Fault_History[1];
        Slab_Fault_History[1] := Slab_Fault_History[0];
        Slab_Fault_History[0] := FaultTimestamp;

        // Activate alarm and start 500 ms hold timer
        faultActive        := TRUE;
        alarmHolding       := TRUE;
        alarmHoldTimer(IN  := TRUE, PT := T#500ms);
    END_IF;

    // -------------------------------------------------------------------------
    // Update alarm state: hold while fault persists or timer running
    // -------------------------------------------------------------------------
    IF faultActive THEN
        // Keep timer running while fault is present
        alarmHoldTimer(IN := TRUE, PT := T#500ms);

        // Alarm stays active while fault or hold timer active
        alarmHolding := THICKNESS_FAULT OR alarmHoldTimer.Q;

        // Release hold tracking once fault clears and timer completes
        IF NOT THICKNESS_FAULT AND alarmHolding AND NOT alarmHoldTimer.Q THEN
            alarmHolding := FALSE;
        END_IF;

        // Clear fault-active flag when fault goes away (hold may continue)
        IF NOT THICKNESS_FAULT THEN
            faultActive := FALSE;
        END_IF;
    END_IF;

    // Final alarm output
    THICKNESS_ALARM := alarmHolding OR faultActive;

    // -------------------------------------------------------------------------
    // Runtime accumulation: only while cutting, signal valid, no fault
    // -------------------------------------------------------------------------
    IF CUTTING_RUN AND NOT THICKNESS_FAULT THEN
        Slab_Runtime_Accumulator := Slab_Runtime_Accumulator + TO_LTIME(CycleTime);
    END_IF;

ELSE
    // Signal invalid: clear alarm and all hold state (PUB001)
    THICKNESS_ALARM  := FALSE;
    alarmHolding     := FALSE;
    faultActive      := FALSE;
    alarmHoldTimer(IN := FALSE);
END_IF;

// ---------------------------------------------------------------------------
// Latch previous scan signal-valid state for edge detection
// ---------------------------------------------------------------------------
signalValidPrev := THICKNESS_SIGNAL_VALID;

END_FUNCTION_BLOCK

(* ---- public-medium-06.patch_base_02.st ---- *)
FUNCTION_BLOCK FB_SlabThicknessMonitor
(*
 * ENGINEERING_CONTRACT
 * =============================================================================
 * Output/State          | Activation          | Retention            | Reset/Deactivation            | Units
 * ----------------------+---------------------+----------------------+-------------------------------+-----------------
 * THICKNESS_ALARM       | Rising edge valid   | Min 500ms hold;      | Signal invalid clears all     | BOOL
 *                       | THICKNESS_FAULT     | continues if fault   | alarm and hold state (PUB001) |
 * Alarm hold timer      | TON(IN: valid &     | TON.ET saturates at  | Signal invalid resets TON     | LTIME (≥500ms)
 *                       |   (fault OR holding))| PT=500ms            |                               |
 * Holding flag          | Fault OR holding    | Self-holds while     | Signal invalid clears         | BOOL
 *                       |                     |   fault OR timer run |                               |
 * Slab_Fault_Counter    | FALSE→TRUE valid    | Accumulates monoton  | None by task spec             | UINT
 *                       | fault transition    | (never auto-reset)   |                               |
 * Slab_Fault_History[0] | New fault entry     | Shifts [n]→[n+1]     | Power-up init to 0            | ARRAY[0..4] DINT
 *                       | writes to index 0   | (0 newest)           |                               |
 * Slab_Runtime_Accumulator| While CUTTING_RUN  | Preserved when       | None by task spec             | LTIME (accumulates)
 *                       | + valid + no fault  | conditions not met   |                               |
 * =============================================================================
 * CONTRACT_RULES [{"kind": "hold_until_reset", "output": "THICKNESS_ALARM", "set_input": "THICKNESS_FAULT", "reset_input": null}]
 *)

VAR_INPUT
    THICKNESS_FAULT        : BOOL;
    THICKNESS_SIGNAL_VALID : BOOL;
    CUTTING_RUN            : BOOL;
    FaultTimestamp         : DINT;
    CycleTime              : TIME;
END_VAR

VAR_OUTPUT
    THICKNESS_ALARM           : BOOL;
    Slab_Fault_Counter        : UINT;
    Slab_Runtime_Accumulator  : LTIME;
    Slab_Fault_History        : ARRAY[0..4] OF DINT;
END_VAR

VAR
    faultRisingEdge    : R_TRIG;
    signalValidPrev    : BOOL;
    alarmHoldTimer     : TON;
    alarmHolding       : BOOL;
    faultActive        : BOOL;
END_VAR

// ---------------------------------------------------------------------------
// Power-up initialization (first scan after instantiation)
// ---------------------------------------------------------------------------
IF NOT alarmHoldTimer.Q AND NOT faultActive AND NOT alarmHolding THEN
    Slab_Fault_Counter       := 0;
    Slab_Runtime_Accumulator := LTIME#0s;
    Slab_Fault_History[0]    := 0;
    Slab_Fault_History[1]    := 0;
    Slab_Fault_History[2]    := 0;
    Slab_Fault_History[3]    := 0;
    Slab_Fault_History[4]    := 0;
END_IF;

// ---------------------------------------------------------------------------
// Detect FALSE→TRUE transition on valid fault signal
// ---------------------------------------------------------------------------
faultRisingEdge(CLK := THICKNESS_FAULT AND THICKNESS_SIGNAL_VALID);

// ---------------------------------------------------------------------------
// Handle signal-valid transitions: clear alarm/hold when signal lost (PUB001)
// ---------------------------------------------------------------------------
IF THICKNESS_SIGNAL_VALID THEN
    IF NOT signalValidPrev THEN
        // Signal just restored after being invalid
        alarmHolding  := FALSE;
        alarmHoldTimer(IN := FALSE);
        faultActive   := FALSE;
    END_IF;

    // -------------------------------------------------------------------------
    // On rising edge of valid fault: record entry and start hold
    // -------------------------------------------------------------------------
    IF faultRisingEdge.Q THEN
        // Increment counter
        Slab_Fault_Counter := Slab_Fault_Counter + UINT#1;

        // Shift history: index 3→4, 2→3, 1→2, 0→1, then write new to 0
        Slab_Fault_History[4] := Slab_Fault_History[3];
        Slab_Fault_History[3] := Slab_Fault_History[2];
        Slab_Fault_History[2] := Slab_Fault_History[1];
        Slab_Fault_History[1] := Slab_Fault_History[0];
        Slab_Fault_History[0] := FaultTimestamp;

        // Activate alarm and start 500 ms hold timer
        faultActive        := TRUE;
        alarmHolding       := TRUE;
        alarmHoldTimer(IN  := TRUE, PT := T#500ms);
    END_IF;

    // -------------------------------------------------------------------------
    // Update alarm state: hold while fault persists or timer running
    // -------------------------------------------------------------------------
    IF faultActive THEN
        // Keep timer running while fault is present
        alarmHoldTimer(IN := TRUE, PT := T#500ms);

        // Alarm stays active while fault or hold timer active
        alarmHolding := THICKNESS_FAULT OR alarmHoldTimer.Q;

        // Release hold tracking once fault clears and timer completes
        IF NOT THICKNESS_FAULT AND alarmHolding AND NOT alarmHoldTimer.Q THEN
            alarmHolding := FALSE;
        END_IF;

        // Clear fault-active flag when fault goes away (hold may continue)
        IF NOT THICKNESS_FAULT THEN
            faultActive := FALSE;
        END_IF;
    END_IF;

    // Final alarm output
    THICKNESS_ALARM := alarmHolding OR faultActive;

    // -------------------------------------------------------------------------
    // Runtime accumulation: only while cutting, signal valid, no fault
    // -------------------------------------------------------------------------
    IF CUTTING_RUN AND NOT THICKNESS_FAULT THEN
        Slab_Runtime_Accumulator := Slab_Runtime_Accumulator + CycleTime;
    END_IF;

ELSE
    // Signal invalid: clear alarm and all hold state (PUB001)
    THICKNESS_ALARM  := FALSE;
    alarmHolding     := FALSE;
    faultActive      := FALSE;
    alarmHoldTimer(IN := FALSE);
END_IF;

// ---------------------------------------------------------------------------
// Latch previous scan signal-valid state for edge detection
// ---------------------------------------------------------------------------
signalValidPrev := THICKNESS_SIGNAL_VALID;

END_FUNCTION_BLOCK

(* ---- public-medium-06.patch_base_03.st ---- *)
FUNCTION_BLOCK FB_SlabThicknessMonitor
(*
 * ENGINEERING_CONTRACT
 * =============================================================================
 * Output/State          | Activation          | Retention            | Reset/Deactivation            | Units
 * ----------------------+---------------------+----------------------+-------------------------------+-----------------
 * THICKNESS_ALARM       | Rising edge valid   | Min 500ms hold;      | Signal invalid clears all     | BOOL
 *                       | THICKNESS_FAULT     | continues if fault   | alarm and hold state (PUB001) |
 * Alarm hold timer      | TON(IN: valid &     | TON.ET saturates at  | Signal invalid resets TON     | LTIME (≥500ms)
 *                       |   (fault OR holding))| PT=500ms            |                               |
 * Holding flag          | Fault OR holding    | Self-holds while     | Signal invalid clears         | BOOL
 *                       |                     |   fault OR timer run |                               |
 * Slab_Fault_Counter    | FALSE→TRUE valid    | Accumulates monoton  | None by task spec             | UINT
 *                       | fault transition    | (never auto-reset)   |                               |
 * Slab_Fault_History[0] | New fault entry     | Shifts [n]→[n+1]     | Power-up init to 0            | ARRAY[0..4] DINT
 *                       | writes to index 0   | (0 newest)           |                               |
 * Slab_Runtime_Accumulator| While CUTTING_RUN  | Preserved when       | None by task spec             | LTIME (accumulates)
 *                       | + valid + no fault  | conditions not met   |                               |
 * =============================================================================
 * CONTRACT_RULES [{"kind": "hold_until_reset", "output": "THICKNESS_ALARM", "set_input": "THICKNESS_FAULT", "reset_input": null}]
 *)

VAR_INPUT
    THICKNESS_FAULT        : BOOL;
    THICKNESS_SIGNAL_VALID : BOOL;
    CUTTING_RUN            : BOOL;
    FaultTimestamp         : DINT;
    CycleTime              : TIME;
END_VAR

VAR_OUTPUT
    THICKNESS_ALARM           : BOOL;
    Slab_Fault_Counter        : UINT;
    Slab_Runtime_Accumulator  : LTIME;
    Slab_Fault_History        : ARRAY[0..4] OF DINT;
END_VAR

VAR
    faultRisingEdge    : R_TRIG;
    signalValidPrev    : BOOL;
    alarmHoldTimer     : TON;
    alarmHolding       : BOOL;
    faultActive        : BOOL;
END_VAR

// ---------------------------------------------------------------------------
// Power-up initialization (first scan after instantiation)
// ---------------------------------------------------------------------------
IF NOT alarmHoldTimer.Q AND NOT faultActive AND NOT alarmHolding THEN
    Slab_Fault_Counter       := 0;
    Slab_Runtime_Accumulator := LTIME#0s;
    Slab_Fault_History[0]    := 0;
    Slab_Fault_History[1]    := 0;
    Slab_Fault_History[2]    := 0;
    Slab_Fault_History[3]    := 0;
    Slab_Fault_History[4]    := 0;
END_IF;

// ---------------------------------------------------------------------------
// Detect FALSE→TRUE transition on valid fault signal
// ---------------------------------------------------------------------------
faultRisingEdge(CLK := THICKNESS_FAULT AND THICKNESS_SIGNAL_VALID);

// ---------------------------------------------------------------------------
// Handle signal-valid transitions: clear alarm/hold when signal lost (PUB001)
// ---------------------------------------------------------------------------
IF THICKNESS_SIGNAL_VALID THEN
    IF NOT signalValidPrev THEN
        // Signal just restored after being invalid
        alarmHolding  := FALSE;
        alarmHoldTimer(IN := FALSE);
        faultActive   := FALSE;
    END_IF;

    // -------------------------------------------------------------------------
    // On rising edge of valid fault: record entry and start hold
    // -------------------------------------------------------------------------
    IF faultRisingEdge.Q THEN
        // Increment counter
        Slab_Fault_Counter := Slab_Fault_Counter + UINT#1;

        // Shift history: index 3→4, 2→3, 1→2, 0→1, then write new to 0
        Slab_Fault_History[4] := Slab_Fault_History[3];
        Slab_Fault_History[3] := Slab_Fault_History[2];
        Slab_Fault_History[2] := Slab_Fault_History[1];
        Slab_Fault_History[1] := Slab_Fault_History[0];
        Slab_Fault_History[0] := FaultTimestamp;

        // Activate alarm and start 500 ms hold timer
        faultActive        := TRUE;
        alarmHolding       := TRUE;
        alarmHoldTimer(IN  := TRUE, PT := T#500ms);
    END_IF;

    // -------------------------------------------------------------------------
    // Update alarm state: hold while fault persists or timer running
    // -------------------------------------------------------------------------
    IF faultActive THEN
        // Keep timer running while fault is present
        alarmHoldTimer(IN := TRUE, PT := T#500ms);

        // Alarm stays active while fault or hold timer active
        alarmHolding := THICKNESS_FAULT OR alarmHoldTimer.Q;

        // Release hold tracking once fault clears and timer completes
        IF NOT THICKNESS_FAULT AND alarmHolding AND NOT alarmHoldTimer.Q THEN
            alarmHolding := FALSE;
        END_IF;

        // Clear fault-active flag when fault goes away (hold may continue)
        IF NOT THICKNESS_FAULT THEN
            faultActive := FALSE;
        END_IF;
    END_IF;

    // Final alarm output
    THICKNESS_ALARM := alarmHolding OR faultActive;

    // -------------------------------------------------------------------------
    // Runtime accumulation: only while cutting, signal valid, no fault
    // -------------------------------------------------------------------------
    IF CUTTING_RUN AND NOT THICKNESS_FAULT THEN
        Slab_Runtime_Accumulator := Slab_Runtime_Accumulator + CycleTime;
    END_IF;

ELSE
    // Signal invalid: clear alarm and all hold state (PUB001)
    THICKNESS_ALARM  := FALSE;
    alarmHolding     := FALSE;
    faultActive      := FALSE;
    alarmHoldTimer(IN := FALSE);
END_IF;

// ---------------------------------------------------------------------------
// Latch previous scan signal-valid state for edge detection
// ---------------------------------------------------------------------------
signalValidPrev := THICKNESS_SIGNAL_VALID;

END_FUNCTION_BLOCK

(* ---- public-medium-06.patch_base_04.st ---- *)
FUNCTION_BLOCK FB_SlabThicknessMonitor
(*
 * ENGINEERING_CONTRACT
 * =============================================================================
 * Output/State          | Activation          | Retention            | Reset/Deactivation            | Units
 * ----------------------+---------------------+----------------------+-------------------------------+-----------------
 * THICKNESS_ALARM       | Rising edge valid   | Min 500ms hold;      | Signal invalid clears all     | BOOL
 *                       | THICKNESS_FAULT     | continues if fault   | alarm and hold state (PUB001) |
 * Alarm hold timer      | TON(IN: valid &     | TON.ET saturates at  | Signal invalid resets TON     | LTIME (≥500ms)
 *                       |   (fault OR holding))| PT=500ms            |                               |
 * Holding flag          | Fault OR holding    | Self-holds while     | Signal invalid clears         | BOOL
 *                       |                     |   fault OR timer run |                               |
 * Slab_Fault_Counter    | FALSE→TRUE valid    | Accumulates monoton  | None by task spec             | UINT
 *                       | fault transition    | (never auto-reset)   |                               |
 * Slab_Fault_History[0] | New fault entry     | Shifts [n]→[n+1]     | Power-up init to 0            | ARRAY[0..4] DINT
 *                       | writes to index 0   | (0 newest)           |                               |
 * Slab_Runtime_Accumulator| While CUTTING_RUN  | Preserved when       | None by task spec             | LTIME (accumulates)
 *                       | + valid + no fault  | conditions not met   |                               |
 * =============================================================================
 * CONTRACT_RULES [{"kind": "hold_until_reset", "output": "THICKNESS_ALARM", "set_input": "THICKNESS_FAULT", "reset_input": null}]
 *)

VAR_INPUT
    THICKNESS_FAULT        : BOOL;
    THICKNESS_SIGNAL_VALID : BOOL;
    CUTTING_RUN            : BOOL;
    FaultTimestamp         : DINT;
    CycleTime              : TIME;
END_VAR

VAR_OUTPUT
    THICKNESS_ALARM           : BOOL;
    Slab_Fault_Counter        : UINT;
    Slab_Runtime_Accumulator  : LTIME;
    Slab_Fault_History        : ARRAY[0..4] OF DINT;
END_VAR

VAR
    faultRisingEdge    : R_TRIG;
    signalValidPrev    : BOOL;
    alarmHoldTimer     : TON;
    alarmHolding       : BOOL;
    faultActive        : BOOL;
END_VAR

// ---------------------------------------------------------------------------
// Power-up initialization (first scan after instantiation)
// ---------------------------------------------------------------------------
IF NOT alarmHoldTimer.Q AND NOT faultActive AND NOT alarmHolding THEN
    Slab_Fault_Counter       := 0;
    Slab_Runtime_Accumulator := LTIME#0ms;
    Slab_Fault_History[0]    := 0;
    Slab_Fault_History[1]    := 0;
    Slab_Fault_History[2]    := 0;
    Slab_Fault_History[3]    := 0;
    Slab_Fault_History[4]    := 0;
END_IF;

// ---------------------------------------------------------------------------
// Detect FALSE→TRUE transition on valid fault signal
// ---------------------------------------------------------------------------
faultRisingEdge(CLK := THICKNESS_FAULT AND THICKNESS_SIGNAL_VALID);

// ---------------------------------------------------------------------------
// Handle signal-valid transitions: clear alarm/hold when signal lost (PUB001)
// ---------------------------------------------------------------------------
IF THICKNESS_SIGNAL_VALID THEN
    IF NOT signalValidPrev THEN
        // Signal just restored after being invalid
        alarmHolding  := FALSE;
        alarmHoldTimer(IN := FALSE);
        faultActive   := FALSE;
    END_IF;

    // -------------------------------------------------------------------------
    // On rising edge of valid fault: record entry and start hold
    // -------------------------------------------------------------------------
    IF faultRisingEdge.Q THEN
        // Increment counter
        Slab_Fault_Counter := Slab_Fault_Counter + UINT#1;

        // Shift history: index 3→4, 2→3, 1→2, 0→1, then write new to 0
        Slab_Fault_History[4] := Slab_Fault_History[3];
        Slab_Fault_History[3] := Slab_Fault_History[2];
        Slab_Fault_History[2] := Slab_Fault_History[1];
        Slab_Fault_History[1] := Slab_Fault_History[0];
        Slab_Fault_History[0] := FaultTimestamp;

        // Activate alarm and start 500 ms hold timer
        faultActive        := TRUE;
        alarmHolding       := TRUE;
        alarmHoldTimer(IN  := TRUE, PT := T#500ms);
    END_IF;

    // -------------------------------------------------------------------------
    // Update alarm state: hold while fault persists or timer running
    // -------------------------------------------------------------------------
    IF faultActive THEN
        // Keep timer running while fault is present
        alarmHoldTimer(IN := TRUE, PT := T#500ms);

        // Alarm stays active while fault or hold timer active
        alarmHolding := THICKNESS_FAULT OR alarmHoldTimer.Q;

        // Release hold tracking once fault clears and timer completes
        IF NOT THICKNESS_FAULT AND alarmHolding AND NOT alarmHoldTimer.Q THEN
            alarmHolding := FALSE;
        END_IF;

        // Clear fault-active flag when fault goes away (hold may continue)
        IF NOT THICKNESS_FAULT THEN
            faultActive := FALSE;
        END_IF;
    END_IF;

    // Final alarm output
    THICKNESS_ALARM := alarmHolding OR faultActive;

    // -------------------------------------------------------------------------
    // Runtime accumulation: only while cutting, signal valid, no fault
    // -------------------------------------------------------------------------
    IF CUTTING_RUN AND NOT THICKNESS_FAULT THEN
        Slab_Runtime_Accumulator := Slab_Runtime_Accumulator + TO_LTIME(CycleTime);
    END_IF;

ELSE
    // Signal invalid: clear alarm and all hold state (PUB001)
    THICKNESS_ALARM  := FALSE;
    alarmHolding     := FALSE;
    faultActive      := FALSE;
    alarmHoldTimer(IN := FALSE);
END_IF;

// ---------------------------------------------------------------------------
// Latch previous scan signal-valid state for edge detection
// ---------------------------------------------------------------------------
signalValidPrev := THICKNESS_SIGNAL_VALID;

END_FUNCTION_BLOCK

(* ---- public-medium-06.raw_candidate_01.st ---- *)
FUNCTION_BLOCK FB_SlabThicknessMonitor
(*
 * ENGINEERING_CONTRACT
 * =============================================================================
 * Output/State          | Activation          | Retention            | Reset/Deactivation            | Units
 * ----------------------+---------------------+----------------------+-------------------------------+-----------------
 * THICKNESS_ALARM       | Rising edge valid   | Min 500ms hold;      | Signal invalid clears all     | BOOL
 *                       | THICKNESS_FAULT     | continues if fault   | alarm and hold state (PUB001) |
 * Alarm hold timer      | TON(IN: valid &     | TON.ET saturates at  | Signal invalid resets TON     | LTIME (≥500ms)
 *                       |   (fault OR holding))| PT=500ms            |                               |
 * Holding flag          | Fault OR holding    | Self-holds while     | Signal invalid clears         | BOOL
 *                       |                     |   fault OR timer run |                               |
 * Slab_Fault_Counter    | FALSE→TRUE valid    | Accumulates monoton  | None by task spec             | UINT
 *                       | fault transition    | (never auto-reset)   |                               |
 * Slab_Fault_History[0] | New fault entry     | Shifts [n]→[n+1]     | Power-up init to 0            | ARRAY[0..4] DINT
 *                       | writes to index 0   | (0 newest)           |                               |
 * Slab_Runtime_Accumulator| While CUTTING_RUN  | Preserved when       | None by task spec             | LTIME (accumulates)
 *                       | + valid + no fault  | conditions not met   |                               |
 * =============================================================================
 * CONTRACT_RULES [{"kind": "hold_until_reset", "output": "THICKNESS_ALARM", "set_input": "THICKNESS_FAULT", "reset_input": null}]
 *)

VAR_INPUT
    THICKNESS_FAULT        : BOOL;
    THICKNESS_SIGNAL_VALID : BOOL;
    CUTTING_RUN            : BOOL;
    FaultTimestamp         : DINT;
    CycleTime              : TIME;
END_VAR

VAR_OUTPUT
    THICKNESS_ALARM           : BOOL;
    Slab_Fault_Counter        : UINT;
    Slab_Runtime_Accumulator  : LTIME;
    Slab_Fault_History        : ARRAY[0..4] OF DINT;
END_VAR

VAR
    faultRisingEdge    : R_TRIG;
    signalValidPrev    : BOOL;
    alarmHoldTimer     : TON;
    alarmHolding       : BOOL;
    faultActive        : BOOL;
END_VAR

// ---------------------------------------------------------------------------
// Power-up initialization (first scan after instantiation)
// ---------------------------------------------------------------------------
IF NOT alarmHoldTimer.Q AND NOT faultActive AND NOT alarmHolding THEN
    Slab_Fault_Counter       := 0;
    Slab_Runtime_Accumulator := LTIME#0s;
    Slab_Fault_History[0]    := 0;
    Slab_Fault_History[1]    := 0;
    Slab_Fault_History[2]    := 0;
    Slab_Fault_History[3]    := 0;
    Slab_Fault_History[4]    := 0;
END_IF

// ---------------------------------------------------------------------------
// Detect FALSE→TRUE transition on valid fault signal
// ---------------------------------------------------------------------------
faultRisingEdge(CLK := THICKNESS_FAULT AND THICKNESS_SIGNAL_VALID);

// ---------------------------------------------------------------------------
// Handle signal-valid transitions: clear alarm/hold when signal lost (PUB001)
// ---------------------------------------------------------------------------
IF THICKNESS_SIGNAL_VALID THEN
    IF NOT signalValidPrev THEN
        // Signal just restored after being invalid
        alarmHolding  := FALSE;
        alarmHoldTimer(IN := FALSE);
        faultActive   := FALSE;
    END_IF

    // -------------------------------------------------------------------------
    // On rising edge of valid fault: record entry and start hold
    // -------------------------------------------------------------------------
    IF faultRisingEdge.Q THEN
        // Increment counter
        Slab_Fault_Counter := Slab_Fault_Counter + UINT#1;

        // Shift history: index 3→4, 2→3, 1→2, 0→1, then write new to 0
        Slab_Fault_History[4] := Slab_Fault_History[3];
        Slab_Fault_History[3] := Slab_Fault_History[2];
        Slab_Fault_History[2] := Slab_Fault_History[1];
        Slab_Fault_History[1] := Slab_Fault_History[0];
        Slab_Fault_History[0] := FaultTimestamp;

        // Activate alarm and start 500 ms hold timer
        faultActive        := TRUE;
        alarmHolding       := TRUE;
        alarmHoldTimer(IN  := TRUE, PT := T#500ms);
    END_IF

    // -------------------------------------------------------------------------
    // Update alarm state: hold while fault persists or timer running
    // -------------------------------------------------------------------------
    IF faultActive THEN
        // Keep timer running while fault is present
        alarmHoldTimer(IN := TRUE, PT := T#500ms);

        // Alarm stays active while fault or hold timer active
        alarmHolding := THICKNESS_FAULT OR alarmHoldTimer.Q;

        // Release hold tracking once fault clears and timer completes
        IF NOT THICKNESS_FAULT AND alarmHolding AND NOT alarmHoldTimer.Q THEN
            alarmHolding := FALSE;
        END_IF;

        // Clear fault-active flag when fault goes away (hold may continue)
        IF NOT THICKNESS_FAULT THEN
            faultActive := FALSE;
        END_IF;
    END_IF;

    // Final alarm output
    THICKNESS_ALARM := alarmHolding OR faultActive;

    // -------------------------------------------------------------------------
    // Runtime accumulation: only while cutting, signal valid, no fault
    // -------------------------------------------------------------------------
    IF CUTTING_RUN AND NOT THICKNESS_FAULT THEN
        Slab_Runtime_Accumulator := Slab_Runtime_Accumulator + CycleTime;
    END_IF;

ELSE
    // Signal invalid: clear alarm and all hold state (PUB001)
    THICKNESS_ALARM  := FALSE;
    alarmHolding     := FALSE;
    faultActive      := FALSE;
    alarmHoldTimer(IN := FALSE);
END_IF;

// ---------------------------------------------------------------------------
// Latch previous scan signal-valid state for edge detection
// ---------------------------------------------------------------------------
signalValidPrev := THICKNESS_SIGNAL_VALID;

END_FUNCTION_BLOCK
